// TIA Portal V21 export
// export: Created 2026-11-10T19:13:02.9074366Z, ExportSetting WithDefaults, DisplayName Totally Integrated Automation Portal, DisplayVersion V21 Update 3, DisplayName STEP 7 Professional, DisplayVersion V21 Update 3, DisplayName STEP 7 Safety, DisplayVersion V21, DisplayName Tech WebApplication, DisplayVersion V21, DisplayName WinCC Basic/Comfort/Advanced, DisplayVersion V21 Update 3, DisplayName WinCC Unified, DisplayVersion V21 Update 3
DATA_BLOCK "DB_TRCV"   // DB13
// stored: AutoNumber true, DBAccessibleFromOPCUA true, DBAccessibleFromWebserver true, InstanceOfName TRCV, OfSystemLibElement TRCV, OfSystemLibVersion 4.0
"TRCV"
   // VAR_INPUT
   //    EN_R : Bool;
   //    ID : CONN_OUC;
   //    LEN : UDInt;
   //    ADHOC : Bool;
   // END_VAR
   // VAR_OUTPUT
   //    NDR : Bool;
   //    BUSY : Bool;
   //    ERROR : Bool;
   //    STATUS : Word;
   //    RCVD_LEN : UDInt;
   // END_VAR
   // VAR_IN_OUT
   //    DATA : Variant;
   //    ADDR : Variant;
   // END_VAR
BEGIN
END_DATA_BLOCK
